(* IEC 61131-3 sources: rusty/tests/lit/single/retain, 3 files *)

(* ---- transitive_fb.st ---- *)
// RUN: %COMPILE %s && %RUN | %CHECK %s
// FB retain members with inline type definitions keep their in-place layout; the
// instances get the retain treatment transitively: the program instance is extracted
// into a retain global, the plain global instance moves to a retain block.
FUNCTION_BLOCK Fb
    VAR RETAIN
        arr : ARRAY[0..2] OF DINT := [1, 2, 3];
        sub : DINT(0..100) := 50;
    END_VAR
END_FUNCTION_BLOCK

PROGRAM mainProg
    VAR
        inst : Fb;
    END_VAR

    inst.arr[0] := inst.arr[0] + 1;
    inst.sub := inst.sub + 1;
END_PROGRAM

VAR_GLOBAL
    gInst : Fb;
END_VAR

FUNCTION main : DINT
    mainProg();
    gInst.arr[2] := 99;
    gInst.sub := gInst.sub + 2;
    printf('%d %d %d$N', mainProg.inst.arr[0], mainProg.inst.arr[1], mainProg.inst.arr[2]); //CHECK: 2 2 3
    printf('%d$N', mainProg.inst.sub);                                                      //CHECK-NEXT: 51
    // Implicitly created global variable backing the program instance
    printf('%d %d$N', __mainProg_inst__retain.arr[0], __mainProg_inst__retain.sub);         //CHECK-NEXT: 2 51
    printf('%d %d$N', gInst.arr[2], gInst.sub);                                             //CHECK-NEXT: 99 52
END_FUNCTION

(* ---- type_shapes.st ---- *)
// RUN: %COMPILE %s && %RUN | %CHECK %s
// Program retain variables with inline type definitions: the extracted inline type
// and the generated retain pointer type must not clash (they both used to be named
// `__<pou>_<var>`), and initializers must land on the generated retain globals.
PROGRAM mainProg
    VAR RETAIN
        arr : ARRAY[0..2] OF DINT := [11, 22, 33];
        sub : DINT(0..100) := 50;
        str : STRING[20] := 'start';
        col : (RED, GREEN, BLUE) := GREEN;
        mat : ARRAY[0..1, 0..2] OF DINT;
        nst : ARRAY[0..1] OF ARRAY[0..2] OF DINT;
        rec : STRUCT a : DINT; b : DINT; END_STRUCT
    END_VAR

    arr[0] := arr[0] + 1;
    sub := sub + 1;
    mat[1, 2] := 42;
    nst[1][2] := 43;
    rec.a := rec.a + 1;
END_PROGRAM

FUNCTION main : DINT
    mainProg();
    printf('%d %d %d$N', mainProg.arr[0], mainProg.arr[1], mainProg.arr[2]); //CHECK: 12 22 33
    printf('%d$N', __mainProg_arr__retain[0]);                               //CHECK-NEXT: 12
    printf('%d %d$N', mainProg.sub, __mainProg_sub__retain);                 //CHECK-NEXT: 51 51
    printf('%s %s$N', REF(mainProg.str), REF(__mainProg_str__retain));       //CHECK-NEXT: start start
    printf('%d %d$N', mainProg.col, __mainProg_col__retain);                 //CHECK-NEXT: 1 1
    printf('%d %d$N', mainProg.mat[1, 2], __mainProg_mat__retain[1, 2]);     //CHECK-NEXT: 42 42
    printf('%d %d$N', mainProg.nst[1][2], __mainProg_nst__retain[1][2]);     //CHECK-NEXT: 43 43
    printf('%d %d$N', mainProg.rec.a, __mainProg_rec__retain.a);             //CHECK-NEXT: 1 1
END_FUNCTION

(* ---- wiring.st ---- *)
// RUN: %COMPILE %s && %RUN | %CHECK %s
VAR_GLOBAL RETAIN
    globalVar : DINT;
END_VAR

PROGRAM mainProg
    VAR RETAIN
        prgVar : DINT;
        prgArr : ARRAY[0..100] OF DINT;
    END_VAR

    prgVar := 20;
    globalVar := 50;
    prgArr[100] := 30;
END_PROGRAM

FUNCTION main : DINT
    mainProg();
    printf('%d$N', mainProg.prgVar); //CHECK: 20
    // Implicitly created global variable
    printf('%d$N', __mainProg_prgVar__retain); //CHECK-NEXT: 20
    printf('%d$N', globalVar); //CHECK-NEXT: 50
    // Variables with an inline type definition get the same treatment
    printf('%d$N', mainProg.prgArr[100]); //CHECK-NEXT: 30
    printf('%d$N', __mainProg_prgArr__retain[100]); //CHECK-NEXT: 30
END_FUNCTION
